Staubli VAL3: loadTRAJ.pgx

public program loadTRAJ(num x_nLib, num& x_nResult)
  local string l_sPath
  local num l_nResult
begin
  if x_nLib>=0
    l_sPath="Disk://data/CustomerLib/lib"+toString("",x_nLib)+"/saveTRAJ"
    //  if libList()
    //    endIf
    x_nResult=trajTemp:libLoad(l_sPath)
    if x_nResult!=0
      popUpMsg("2")
      call rs:setAlarm(300,0)
    endIf
  else
    call rs:setAlarm(302,0)
  endIf
end
